Fanuc KAREL source: compact_preamble.KL

PROGRAM KB00008
%NOLOCKGROUP
VAR
P1:REAL;RESULT:REAL
BEGIN
P1=1.0
RESULT=ASIN(P1)
END KB00008
